(* IEC 61131-3 sources: safety-mesh/modules/plc/DUTs, 2 files *)

(* ---- ST_RobotDH.st ---- *)
// Denavit-Hartenberg parameters
// Index 0..5 = joints A1..A6, same order as ST_RobotPose.aJoints.
TYPE ST_RobotDH :
STRUCT
    nJointCount   : USINT;                // number of valid joints
    aA_m          : ARRAY[0..5] OF LREAL; // link length a [m]
    aAlpha_deg    : ARRAY[0..5] OF LREAL; // link twist alpha [deg]
    aD_m          : ARRAY[0..5] OF LREAL; // link offset d [m]
    aThetaOff_deg : ARRAY[0..5] OF LREAL; // joint angle offset theta [deg]
    aMin_deg      : ARRAY[0..5] OF LREAL; // lower joint limit [deg]
    aMax_deg      : ARRAY[0..5] OF LREAL; // upper joint limit [deg]
END_STRUCT
END_TYPE

(* ---- ST_RobotPose.st ---- *)
TYPE ST_RobotPose :
STRUCT
    nCycle   : UDINT;            // incremented every write → detects stale data
    nJointCount : USINT;         // number of valid entries in aJoints
    fTcpX, fTcpY, fTcpZ : LREAL; // cartesian coordinates of TCP in robot frame
    fTcpA, fTcpB, fTcpC : LREAL; // orientation
    aJoints  : ARRAY[0..5] OF LREAL;
END_STRUCT
END_TYPE
